FUNCTION_BLOCK fbHome
VAR
	LivingRoom : fbRoomLiving;
END_VAR

LivingRoom();

END_FUNCTION_BLOCK

(* stored: Version 1.1.0.1
   POU fbHome: Id {d86ccfb6-79d9-4713-bab4-002d4cb6edd7}, SpecialFunc None *)
